(* IEC 61131-3 sources: trust-platform/conformance/cases/strings/cfm_strings_slice_concat_001, 1 file *)

(* ---- program.st ---- *)
PROGRAM Main
VAR
    text : STRING[16] := 'ABCD';
    second : CHAR := ' ';
    length : INT := INT#0;
    combined : STRING[16] := '';
END_VAR

second := text[2];
length := LEN(text);
combined := CONCAT(text, 'EF');
END_PROGRAM
